TYPE E_CamErrorSource :
(
    CAM_SOURCE_NONE := 0,
    CAM_SOURCE_RECIPE,
    CAM_SOURCE_MASTER_AXIS,
    CAM_SOURCE_SLAVE_AXIS,
    CAM_SOURCE_TABLE_LOAD,
    CAM_SOURCE_TABLE_CHARACTERISTICS,
    CAM_SOURCE_CAM_IN,
    CAM_SOURCE_CAM_OUT
);
END_TYPE

(* stored: Version 1.1.0.1, ProductVersion 3.1.4024.16
   DUT E_CamErrorSource: Id {f93adb1f-408f-4e40-b084-b60ac4754ef9} *)
